FUNCTION_BLOCK basicSubestacao (* Logica unica do QGBT da Subestacao: Masterpact, fonte das barras, planta nos geradores e cargas liberadas *)
  (* Standard: 61499-2 *)
  (* Version 1.3, 04/11/2026, Hidryco, Hidryco, 1.3: comandos do legado REQ_ABRIR_/REQ_FECHAR_1Qx (hmiAbrir/hmiFechar1qx TRUE = mesmo comando do hmiCmdDisjuntor, mesmas permissoes e pulso; FALSE nao faz nada). 1.2: anel - disjuntor com fechamento pendente conta como fechado e o pulso de fechar e cortado se o anel deixar de ter um aberto (nunca as duas QTAM em paralelo). 1.1: comandos de abrir/fechar dos Masterpact 1Q1/1Q0/1Q2 com intertravamentos e aviso de sem resposta; reservas no unifilar. 1.0: QGBT 440 V com 2 QTAM (AGC 150), 1Q1/1Q0/1Q2 e cargas liberadas no gerador *)
  PACKAGE Hidryco.HidrycoLib;
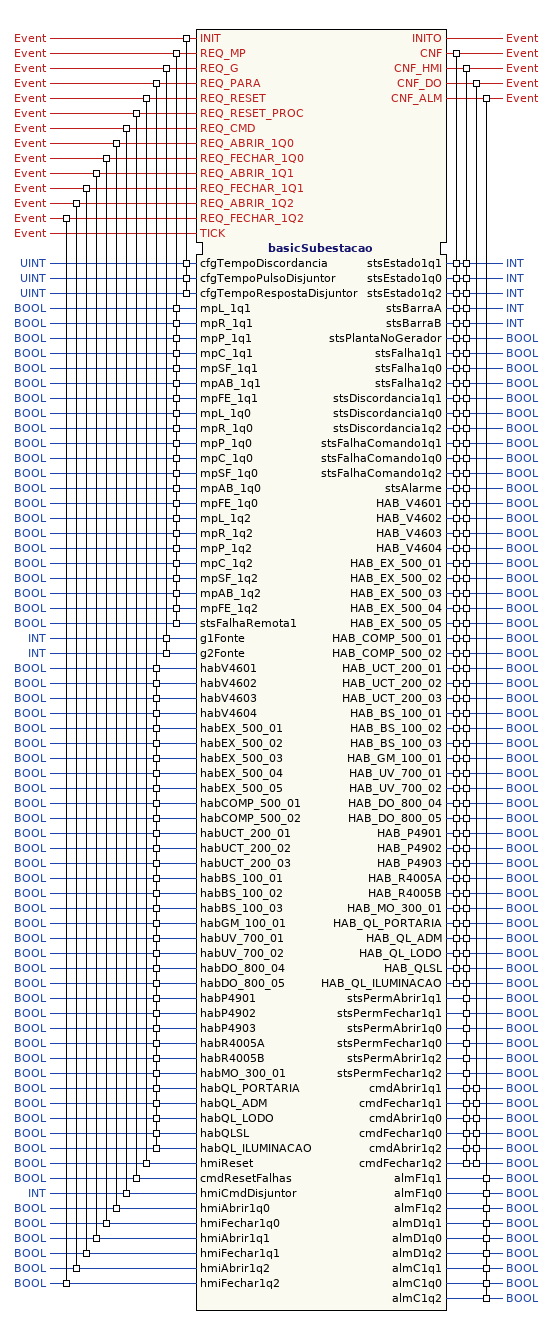
  EVENT_INPUT
    INIT WITH cfgTempoDiscordancia, cfgTempoPulsoDisjuntor, cfgTempoRespostaDisjuntor; (* Inicializacao *)
    REQ_MP WITH mpL_1q1, mpR_1q1, mpP_1q1, mpC_1q1, mpSF_1q1, mpAB_1q1, mpFE_1q1, mpL_1q0, mpR_1q0, mpP_1q0, mpC_1q0, mpSF_1q0, mpAB_1q0, mpFE_1q0, mpL_1q2, mpR_1q2, mpP_1q2, mpC_1q2, mpSF_1q2, mpAB_1q2, mpFE_1q2, stsFalhaRemota1; (* Sinais dos Masterpact e da remota 1 *)
    REQ_G WITH g1Fonte, g2Fonte; (* Estado das QTAM (geradores) *)
    REQ_PARA WITH habV4601, habV4602, habV4603, habV4604, habEX_500_01, habEX_500_02, habEX_500_03, habEX_500_04, habEX_500_05, habCOMP_500_01, habCOMP_500_02, habUCT_200_01, habUCT_200_02, habUCT_200_03, habBS_100_01, habBS_100_02, habBS_100_03, habGM_100_01, habUV_700_01, habUV_700_02, habDO_800_04, habDO_800_05, habP4901, habP4902, habP4903, habR4005A, habR4005B, habMO_300_01, habQL_PORTARIA, habQL_ADM, habQL_LODO, habQLSL, habQL_ILUMINACAO; (* Cargas liberadas no gerador (persistentes) *)
    REQ_RESET WITH hmiReset; (* Reconhecimento pela IHM *)
    REQ_RESET_PROC WITH cmdResetFalhas; (* Reconhecimento pelo processo *)
    REQ_CMD WITH hmiCmdDisjuntor; (* Comando da IHM para os Masterpact *)
    REQ_ABRIR_1Q0 WITH hmiAbrir1q0; (* IHM (legado): ABRIR_1Q0 *)
    REQ_FECHAR_1Q0 WITH hmiFechar1q0; (* IHM (legado): FECHAR_1Q0 *)
    REQ_ABRIR_1Q1 WITH hmiAbrir1q1; (* IHM (legado): ABRIR_1Q1 *)
    REQ_FECHAR_1Q1 WITH hmiFechar1q1; (* IHM (legado): FECHAR_1Q1 *)
    REQ_ABRIR_1Q2 WITH hmiAbrir1q2; (* IHM (legado): ABRIR_1Q2 *)
    REQ_FECHAR_1Q2 WITH hmiFechar1q2; (* IHM (legado): FECHAR_1Q2 *)
    TICK; (* Base de tempo de 1 s *)
  END_EVENT
  EVENT_OUTPUT
    INITO; (* Inicializacao concluida *)
    CNF WITH stsEstado1q1, stsEstado1q0, stsEstado1q2, stsBarraA, stsBarraB, stsPlantaNoGerador, stsFalha1q1, stsFalha1q0, stsFalha1q2, stsDiscordancia1q1, stsDiscordancia1q0, stsDiscordancia1q2, stsFalhaComando1q1, stsFalhaComando1q0, stsFalhaComando1q2, stsAlarme, HAB_V4601, HAB_V4602, HAB_V4603, HAB_V4604, HAB_EX_500_01, HAB_EX_500_02, HAB_EX_500_03, HAB_EX_500_04, HAB_EX_500_05, HAB_COMP_500_01, HAB_COMP_500_02, HAB_UCT_200_01, HAB_UCT_200_02, HAB_UCT_200_03, HAB_BS_100_01, HAB_BS_100_02, HAB_BS_100_03, HAB_GM_100_01, HAB_UV_700_01, HAB_UV_700_02, HAB_DO_800_04, HAB_DO_800_05, HAB_P4901, HAB_P4902, HAB_P4903, HAB_R4005A, HAB_R4005B, HAB_MO_300_01, HAB_QL_PORTARIA, HAB_QL_ADM, HAB_QL_LODO, HAB_QLSL, HAB_QL_ILUMINACAO; (* Estados e cargas liberadas (na mudanca) *)
    CNF_HMI WITH stsEstado1q1, stsEstado1q0, stsEstado1q2, stsBarraA, stsBarraB, stsPlantaNoGerador, stsFalha1q1, stsFalha1q0, stsFalha1q2, stsDiscordancia1q1, stsDiscordancia1q0, stsDiscordancia1q2, stsFalhaComando1q1, stsFalhaComando1q0, stsFalhaComando1q2, stsAlarme, HAB_V4601, HAB_V4602, HAB_V4603, HAB_V4604, HAB_EX_500_01, HAB_EX_500_02, HAB_EX_500_03, HAB_EX_500_04, HAB_EX_500_05, HAB_COMP_500_01, HAB_COMP_500_02, HAB_UCT_200_01, HAB_UCT_200_02, HAB_UCT_200_03, HAB_BS_100_01, HAB_BS_100_02, HAB_BS_100_03, HAB_GM_100_01, HAB_UV_700_01, HAB_UV_700_02, HAB_DO_800_04, HAB_DO_800_05, HAB_P4901, HAB_P4902, HAB_P4903, HAB_R4005A, HAB_R4005B, HAB_MO_300_01, HAB_QL_PORTARIA, HAB_QL_ADM, HAB_QL_LODO, HAB_QLSL, HAB_QL_ILUMINACAO, stsPermAbrir1q1, stsPermFechar1q1, stsPermAbrir1q0, stsPermFechar1q0, stsPermAbrir1q2, stsPermFechar1q2, cmdAbrir1q1, cmdFechar1q1, cmdAbrir1q0, cmdFechar1q0, cmdAbrir1q2, cmdFechar1q2; (* Status para a IHM (na mudanca) *)
    CNF_DO WITH cmdAbrir1q1, cmdFechar1q1, cmdAbrir1q0, cmdFechar1q0, cmdAbrir1q2, cmdFechar1q2; (* Comandos dos Masterpact para o A8 da remota 1 (na mudanca) *)
    CNF_ALM WITH almF1q1, almF1q0, almF1q2, almD1q1, almD1q0, almD1q2, almC1q1, almC1q0, almC1q2; (* Alarmes para os ALARM_BIT (na mudanca) *)
  END_EVENT
  VAR_INPUT
    cfgTempoDiscordancia : UINT := 5; (* Tempo (s) com aberto/fechado discordantes para o aviso de posicao indefinida *)
    cfgTempoPulsoDisjuntor : UINT := 1; (* Tempo (s) do pulso de abrir/fechar dos Masterpact (o pulso acaba antes se o disjuntor mudar de estado) *)
    cfgTempoRespostaDisjuntor : UINT := 5; (* Tempo (s) para o Masterpact mudar de estado depois do comando (senao: aviso de sem resposta) *)
    mpL_1q1 : BOOL; (* Local 1Q1 *)
    mpR_1q1 : BOOL; (* Remoto 1Q1 *)
    mpP_1q1 : BOOL; (* Pronto para fechar 1Q1 *)
    mpC_1q1 : BOOL; (* Mola carregada 1Q1 *)
    mpSF_1q1 : BOOL; (* Sem falha 1Q1 *)
    mpAB_1q1 : BOOL; (* Aberto 1Q1 *)
    mpFE_1q1 : BOOL; (* Fechado 1Q1 *)
    mpL_1q0 : BOOL; (* Local 1Q0 *)
    mpR_1q0 : BOOL; (* Remoto 1Q0 *)
    mpP_1q0 : BOOL; (* Pronto para fechar 1Q0 *)
    mpC_1q0 : BOOL; (* Mola carregada 1Q0 *)
    mpSF_1q0 : BOOL; (* Sem falha 1Q0 *)
    mpAB_1q0 : BOOL; (* Aberto 1Q0 *)
    mpFE_1q0 : BOOL; (* Fechado 1Q0 *)
    mpL_1q2 : BOOL; (* Local 1Q2 *)
    mpR_1q2 : BOOL; (* Remoto 1Q2 *)
    mpP_1q2 : BOOL; (* Pronto para fechar 1Q2 *)
    mpC_1q2 : BOOL; (* Mola carregada 1Q2 *)
    mpSF_1q2 : BOOL; (* Sem falha 1Q2 *)
    mpAB_1q2 : BOOL; (* Aberto 1Q2 *)
    mpFE_1q2 : BOOL; (* Fechado 1Q2 *)
    stsFalhaRemota1 : BOOL; (* Falha de comunicacao com a remota 1 *)
    g1Fonte : INT; (* G1 (QTAM 2): fonte da saida (0 sem, 1 rede, 2 gerador, 3 indefinida) *)
    g2Fonte : INT; (* G2 (QTAM 1): fonte da saida *)
    habV4601 : BOOL; (* IHM: V4601 - Soprador 01 liberado no gerador *)
    habV4602 : BOOL; (* IHM: V4602 - Soprador 02 liberado no gerador *)
    habV4603 : BOOL; (* IHM: V4603 - Soprador 03 liberado no gerador *)
    habV4604 : BOOL; (* IHM: V4604 - Soprador 04 liberado no gerador *)
    habEX_500_01 : BOOL; (* IHM: 500-EX-01 - Exaustor 01 liberado no gerador *)
    habEX_500_02 : BOOL; (* IHM: 500-EX-02 - Exaustor 02 liberado no gerador *)
    habEX_500_03 : BOOL; (* IHM: 500-EX-03 - Exaustor 03 liberado no gerador *)
    habEX_500_04 : BOOL; (* IHM: 500-EX-04 - Exaustor 04 liberado no gerador *)
    habEX_500_05 : BOOL; (* IHM: 500-EX-05 - Exaustor 05 liberado no gerador *)
    habCOMP_500_01 : BOOL; (* IHM: 500-COMP-01 - Compressor 01 liberado no gerador *)
    habCOMP_500_02 : BOOL; (* IHM: 500-COMP-02 - Compressor 02 liberado no gerador *)
    habUCT_200_01 : BOOL; (* IHM: 200-UCT-01 - Unid. compacta 01 liberado no gerador *)
    habUCT_200_02 : BOOL; (* IHM: 200-UCT-02 - Unid. compacta 02 liberado no gerador *)
    habUCT_200_03 : BOOL; (* IHM: 200-UCT-03 - Unid. compacta 03 liberado no gerador *)
    habBS_100_01 : BOOL; (* IHM: 100-BS-01 - Bomba 01 liberado no gerador *)
    habBS_100_02 : BOOL; (* IHM: 100-BS-02 - Bomba 02 liberado no gerador *)
    habBS_100_03 : BOOL; (* IHM: 100-BS-03 - Bomba 03 liberado no gerador *)
    habGM_100_01 : BOOL; (* IHM: 100-GM-01 - Grade mecanizada liberado no gerador *)
    habUV_700_01 : BOOL; (* IHM: 700-UV-01 - Sistema UV 01 liberado no gerador *)
    habUV_700_02 : BOOL; (* IHM: 700-UV-02 - Sistema UV 02 liberado no gerador *)
    habDO_800_04 : BOOL; (* IHM: 800-DO-04 - Bomba dosadora 04 liberado no gerador *)
    habDO_800_05 : BOOL; (* IHM: 800-DO-05 - Bomba dosadora 05 liberado no gerador *)
    habP4901 : BOOL; (* IHM: P4901 - Bomba submersível 01 liberado no gerador *)
    habP4902 : BOOL; (* IHM: P4902 - Bomba submersível 02 liberado no gerador *)
    habP4903 : BOOL; (* IHM: P4903 - Bomba submersível 03 liberado no gerador *)
    habR4005A : BOOL; (* IHM: R4005A - Bomba horizontal A liberado no gerador *)
    habR4005B : BOOL; (* IHM: R4005B - Bomba horizontal B liberado no gerador *)
    habMO_300_01 : BOOL; (* IHM: 300-MO-01 - Misturador 01 liberado no gerador *)
    habQL_PORTARIA : BOOL; (* IHM: QL Portaria liberado no gerador *)
    habQL_ADM : BOOL; (* IHM: QL Administração liberado no gerador *)
    habQL_LODO : BOOL; (* IHM: QL Lodo liberado no gerador *)
    habQLSL : BOOL; (* IHM: QL Sala de quadros liberado no gerador *)
    habQL_ILUMINACAO : BOOL; (* IHM: QL Iluminação externa liberado no gerador *)
    hmiReset : BOOL; (* IHM: reconhecimento *)
    cmdResetFalhas : BOOL; (* Processo: reconhecimento (com E_RESET_FALHAS) *)
    hmiCmdDisjuntor : INT; (* IHM: 1 abrir 1Q1, 2 fechar 1Q1, 3 abrir 1Q0, 4 fechar 1Q0, 5 abrir 1Q2, 6 fechar 1Q2 *)
    hmiAbrir1q0 : BOOL; (* IHM (legado): ABRIR_1Q0, TRUE = executa *)
    hmiFechar1q0 : BOOL; (* IHM (legado): FECHAR_1Q0, TRUE = executa *)
    hmiAbrir1q1 : BOOL; (* IHM (legado): ABRIR_1Q1, TRUE = executa *)
    hmiFechar1q1 : BOOL; (* IHM (legado): FECHAR_1Q1, TRUE = executa *)
    hmiAbrir1q2 : BOOL; (* IHM (legado): ABRIR_1Q2, TRUE = executa *)
    hmiFechar1q2 : BOOL; (* IHM (legado): FECHAR_1Q2, TRUE = executa *)
  END_VAR
  VAR_OUTPUT
    stsEstado1q1 : INT; (* Disjuntor 1Q1: 0 indefinido (sem comunicacao), 1 aberto, 2 fechado, 3 discordante *)
    stsEstado1q0 : INT; (* Disjuntor 1Q0: 0 indefinido (sem comunicacao), 1 aberto, 2 fechado, 3 discordante *)
    stsEstado1q2 : INT; (* Disjuntor 1Q2: 0 indefinido (sem comunicacao), 1 aberto, 2 fechado, 3 discordante *)
    stsBarraA : INT; (* Fonte da barra A (1Q1): 0 sem alimentacao, 1 rede, 2 gerador, 3 indefinida *)
    stsBarraB : INT; (* Fonte da barra B (1Q2): 0 sem alimentacao, 1 rede, 2 gerador, 3 indefinida *)
    stsPlantaNoGerador : BOOL; (* Alguma QTAM com o disjuntor do gerador fechado (planta nos geradores) *)
    stsFalha1q1 : BOOL; (* Disjuntor 1Q1 em falha (desarmado) *)
    stsFalha1q0 : BOOL; (* Disjuntor 1Q0 em falha (desarmado) *)
    stsFalha1q2 : BOOL; (* Disjuntor 1Q2 em falha (desarmado) *)
    stsDiscordancia1q1 : BOOL; (* Disjuntor 1Q1: posição indefinida (aberto e fechado discordantes) *)
    stsDiscordancia1q0 : BOOL; (* Disjuntor 1Q0: posição indefinida (aberto e fechado discordantes) *)
    stsDiscordancia1q2 : BOOL; (* Disjuntor 1Q2: posição indefinida (aberto e fechado discordantes) *)
    stsFalhaComando1q1 : BOOL; (* Disjuntor 1Q1 não respondeu ao comando de abrir/fechar *)
    stsFalhaComando1q0 : BOOL; (* Disjuntor 1Q0 não respondeu ao comando de abrir/fechar *)
    stsFalhaComando1q2 : BOOL; (* Disjuntor 1Q2 não respondeu ao comando de abrir/fechar *)
    stsAlarme : BOOL; (* Algum alarme do QGBT *)
    HAB_V4601 : BOOL; (* V4601 - Soprador 01 liberado para operar com a planta nos geradores *)
    HAB_V4602 : BOOL; (* V4602 - Soprador 02 liberado para operar com a planta nos geradores *)
    HAB_V4603 : BOOL; (* V4603 - Soprador 03 liberado para operar com a planta nos geradores *)
    HAB_V4604 : BOOL; (* V4604 - Soprador 04 liberado para operar com a planta nos geradores *)
    HAB_EX_500_01 : BOOL; (* 500-EX-01 - Exaustor 01 liberado para operar com a planta nos geradores *)
    HAB_EX_500_02 : BOOL; (* 500-EX-02 - Exaustor 02 liberado para operar com a planta nos geradores *)
    HAB_EX_500_03 : BOOL; (* 500-EX-03 - Exaustor 03 liberado para operar com a planta nos geradores *)
    HAB_EX_500_04 : BOOL; (* 500-EX-04 - Exaustor 04 liberado para operar com a planta nos geradores *)
    HAB_EX_500_05 : BOOL; (* 500-EX-05 - Exaustor 05 liberado para operar com a planta nos geradores *)
    HAB_COMP_500_01 : BOOL; (* 500-COMP-01 - Compressor 01 liberado para operar com a planta nos geradores *)
    HAB_COMP_500_02 : BOOL; (* 500-COMP-02 - Compressor 02 liberado para operar com a planta nos geradores *)
    HAB_UCT_200_01 : BOOL; (* 200-UCT-01 - Unid. compacta 01 liberado para operar com a planta nos geradores *)
    HAB_UCT_200_02 : BOOL; (* 200-UCT-02 - Unid. compacta 02 liberado para operar com a planta nos geradores *)
    HAB_UCT_200_03 : BOOL; (* 200-UCT-03 - Unid. compacta 03 liberado para operar com a planta nos geradores *)
    HAB_BS_100_01 : BOOL; (* 100-BS-01 - Bomba 01 liberado para operar com a planta nos geradores *)
    HAB_BS_100_02 : BOOL; (* 100-BS-02 - Bomba 02 liberado para operar com a planta nos geradores *)
    HAB_BS_100_03 : BOOL; (* 100-BS-03 - Bomba 03 liberado para operar com a planta nos geradores *)
    HAB_GM_100_01 : BOOL; (* 100-GM-01 - Grade mecanizada liberado para operar com a planta nos geradores *)
    HAB_UV_700_01 : BOOL; (* 700-UV-01 - Sistema UV 01 liberado para operar com a planta nos geradores *)
    HAB_UV_700_02 : BOOL; (* 700-UV-02 - Sistema UV 02 liberado para operar com a planta nos geradores *)
    HAB_DO_800_04 : BOOL; (* 800-DO-04 - Bomba dosadora 04 liberado para operar com a planta nos geradores *)
    HAB_DO_800_05 : BOOL; (* 800-DO-05 - Bomba dosadora 05 liberado para operar com a planta nos geradores *)
    HAB_P4901 : BOOL; (* P4901 - Bomba submersível 01 liberado para operar com a planta nos geradores *)
    HAB_P4902 : BOOL; (* P4902 - Bomba submersível 02 liberado para operar com a planta nos geradores *)
    HAB_P4903 : BOOL; (* P4903 - Bomba submersível 03 liberado para operar com a planta nos geradores *)
    HAB_R4005A : BOOL; (* R4005A - Bomba horizontal A liberado para operar com a planta nos geradores *)
    HAB_R4005B : BOOL; (* R4005B - Bomba horizontal B liberado para operar com a planta nos geradores *)
    HAB_MO_300_01 : BOOL; (* 300-MO-01 - Misturador 01 liberado para operar com a planta nos geradores *)
    HAB_QL_PORTARIA : BOOL; (* QL Portaria liberado para operar com a planta nos geradores *)
    HAB_QL_ADM : BOOL; (* QL Administração liberado para operar com a planta nos geradores *)
    HAB_QL_LODO : BOOL; (* QL Lodo liberado para operar com a planta nos geradores *)
    HAB_QLSL : BOOL; (* QL Sala de quadros liberado para operar com a planta nos geradores *)
    HAB_QL_ILUMINACAO : BOOL; (* QL Iluminação externa liberado para operar com a planta nos geradores *)
    stsPermAbrir1q1 : BOOL; (* IHM: abrir o 1Q1 permitido *)
    stsPermFechar1q1 : BOOL; (* IHM: fechar o 1Q1 permitido *)
    stsPermAbrir1q0 : BOOL; (* IHM: abrir o 1Q0 permitido *)
    stsPermFechar1q0 : BOOL; (* IHM: fechar o 1Q0 permitido *)
    stsPermAbrir1q2 : BOOL; (* IHM: abrir o 1Q2 permitido *)
    stsPermFechar1q2 : BOOL; (* IHM: fechar o 1Q2 permitido *)
    cmdAbrir1q1 : BOOL; (* Pulso de abrir o 1Q1 (bobina MX) *)
    cmdFechar1q1 : BOOL; (* Pulso de fechar o 1Q1 (bobina XF) *)
    cmdAbrir1q0 : BOOL; (* Pulso de abrir o 1Q0 (bobina MX) *)
    cmdFechar1q0 : BOOL; (* Pulso de fechar o 1Q0 (bobina XF) *)
    cmdAbrir1q2 : BOOL; (* Pulso de abrir o 1Q2 (bobina MX) *)
    cmdFechar1q2 : BOOL; (* Pulso de fechar o 1Q2 (bobina XF) *)
    almF1q1 : BOOL; (* ALARM_BIT Disjuntor 1Q1 em falha (desarmado) *)
    almF1q0 : BOOL; (* ALARM_BIT Disjuntor 1Q0 em falha (desarmado) *)
    almF1q2 : BOOL; (* ALARM_BIT Disjuntor 1Q2 em falha (desarmado) *)
    almD1q1 : BOOL; (* ALARM_BIT Disjuntor 1Q1: posição indefinida (aberto e fechado discordantes) *)
    almD1q0 : BOOL; (* ALARM_BIT Disjuntor 1Q0: posição indefinida (aberto e fechado discordantes) *)
    almD1q2 : BOOL; (* ALARM_BIT Disjuntor 1Q2: posição indefinida (aberto e fechado discordantes) *)
    almC1q1 : BOOL; (* ALARM_BIT Disjuntor 1Q1 não respondeu ao comando de abrir/fechar *)
    almC1q0 : BOOL; (* ALARM_BIT Disjuntor 1Q0 não respondeu ao comando de abrir/fechar *)
    almC1q2 : BOOL; (* ALARM_BIT Disjuntor 1Q2 não respondeu ao comando de abrir/fechar *)
  END_VAR
  VAR
    cmdDj : INT; (* Comando do disjuntor deste ciclo (hmiCmdDisjuntor ou comando do legado) *)
    initDone : BOOL;
    initPass : BOOL;
    bMudou : BOOL;
    u1q1 : UDINT; (* Segundos com aberto/fechado discordantes *)
    u1q0 : UDINT; (* Segundos com aberto/fechado discordantes *)
    u1q2 : UDINT; (* Segundos com aberto/fechado discordantes *)
    e1q1 : INT;
    e1q0 : INT;
    e1q2 : INT;
    wSts : DWORD;
    oldSts : DWORD := 16#FFFFFFFF;
    wHab : DWORD;
    oldHab : DWORD := 16#FFFFFFFF;
    wHab2 : DWORD;
    oldHab2 : DWORD := 16#FFFFFFFF;
    wAlm : WORD;
    oldAlm : WORD := 16#FFFF;
    wPerm : WORD;
    oldPerm : WORD := 16#FFFF;
    wDo : WORD;
    oldDo : WORD := 16#FFFF;
    o_stsEstado1q1 : INT := -1;
    o_stsEstado1q0 : INT := -1;
    o_stsEstado1q2 : INT := -1;
    o_stsBarraA : INT := -1;
    o_stsBarraB : INT := -1;
    tA1q1 : UINT; (* Pulso de abrir restante (s) *)
    tF1q1 : UINT; (* Pulso de fechar restante (s) *)
    uR1q1 : UINT; (* Tempo restante para a resposta (s) *)
    tA1q0 : UINT; (* Pulso de abrir restante (s) *)
    tF1q0 : UINT; (* Pulso de fechar restante (s) *)
    uR1q0 : UINT; (* Tempo restante para a resposta (s) *)
    tA1q2 : UINT; (* Pulso de abrir restante (s) *)
    tF1q2 : UINT; (* Pulso de fechar restante (s) *)
    uR1q2 : UINT; (* Tempo restante para a resposta (s) *)
    alvo1q1 : INT; (* Estado esperado depois do comando (0 nenhum, 1 aberto, 2 fechado) *)
    alvo1q0 : INT; (* Estado esperado depois do comando (0 nenhum, 1 aberto, 2 fechado) *)
    alvo1q2 : INT; (* Estado esperado depois do comando (0 nenhum, 1 aberto, 2 fechado) *)
  END_VAR
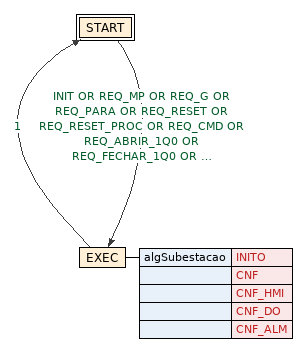
  EC_STATES
    START; (* Estado inicial *)
    EXEC : algSubestacao -> INITO, -> CNF, -> CNF_HMI, -> CNF_DO, -> CNF_ALM; (* Executa a logica; o algoritmo decide quais eventos saem *)
  END_STATES
  EC_TRANSITIONS
    START TO EXEC := INIT OR REQ_MP OR REQ_G OR REQ_PARA OR REQ_RESET OR REQ_RESET_PROC OR REQ_CMD OR REQ_ABRIR_1Q0 OR REQ_FECHAR_1Q0 OR REQ_ABRIR_1Q1 OR REQ_FECHAR_1Q1 OR REQ_ABRIR_1Q2 OR REQ_FECHAR_1Q2 OR TICK;
    EXEC TO START := 1;
  END_TRANSITIONS
  ALGORITHM algSubestacao IN ST: (* Logica completa do QGBT (um unico algoritmo) *)
(* =====================================================================
   basicSubestacao v1.1 - QGBT 440 V da ETE Tijuco Preto
   QTAM 1 (G2) -> 1Q1 -> barra A; QTAM 2 (G1) -> 1Q2 -> barra B; 1Q0 acopla.
   - Masterpact: 2 fechado, 1 aberto, 3 aberto/fechado discordantes,
     0 indefinido (remota 1 sem comunicacao); aviso de discordancia apos
     cfgTempoDiscordancia s; alarme de falha com "sem falha" = FALSE;
   - fonte de cada barra pelo seu Masterpact ou pelo acoplamento 1Q0;
   - planta nos geradores = alguma QTAM com o disjuntor do gerador fechado
     (vale mesmo com a remota 1 sem comunicacao);
   - cargas liberadas no gerador: escolha do operador (persistente), saidas
     HAB_* para os CATs de processo (geradorHabilita);
   - v1.1: comandos de abrir/fechar dos Masterpact com intertravamentos.
   ===================================================================== *)

INITO   := FALSE;
CNF     := FALSE;
CNF_HMI := FALSE;
CNF_DO  := FALSE;
CNF_ALM := FALSE;
IF INIT THEN
    initDone := TRUE;
    initPass := TRUE;
    INITO    := TRUE;
END_IF;
IF NOT initDone THEN
    RETURN;
END_IF;

(* ---- 1Q1 ---- *)
IF stsFalhaRemota1 THEN
    e1q1 := 0;
ELSIF mpAB_1q1 AND NOT mpFE_1q1 THEN
    e1q1 := 1;
ELSIF mpFE_1q1 AND NOT mpAB_1q1 THEN
    e1q1 := 2;
ELSE
    e1q1 := 3;
END_IF;
IF e1q1 = 3 THEN
    IF TICK AND u1q1 < UINT_TO_UDINT(cfgTempoDiscordancia) THEN
        u1q1 := u1q1 + 1;
    END_IF;
ELSE
    u1q1 := 0;
END_IF;
stsEstado1q1 := e1q1;
stsDiscordancia1q1 := e1q1 = 3 AND u1q1 >= UINT_TO_UDINT(cfgTempoDiscordancia);
stsFalha1q1 := NOT stsFalhaRemota1 AND NOT mpSF_1q1;

(* ---- 1Q0 ---- *)
IF stsFalhaRemota1 THEN
    e1q0 := 0;
ELSIF mpAB_1q0 AND NOT mpFE_1q0 THEN
    e1q0 := 1;
ELSIF mpFE_1q0 AND NOT mpAB_1q0 THEN
    e1q0 := 2;
ELSE
    e1q0 := 3;
END_IF;
IF e1q0 = 3 THEN
    IF TICK AND u1q0 < UINT_TO_UDINT(cfgTempoDiscordancia) THEN
        u1q0 := u1q0 + 1;
    END_IF;
ELSE
    u1q0 := 0;
END_IF;
stsEstado1q0 := e1q0;
stsDiscordancia1q0 := e1q0 = 3 AND u1q0 >= UINT_TO_UDINT(cfgTempoDiscordancia);
stsFalha1q0 := NOT stsFalhaRemota1 AND NOT mpSF_1q0;

(* ---- 1Q2 ---- *)
IF stsFalhaRemota1 THEN
    e1q2 := 0;
ELSIF mpAB_1q2 AND NOT mpFE_1q2 THEN
    e1q2 := 1;
ELSIF mpFE_1q2 AND NOT mpAB_1q2 THEN
    e1q2 := 2;
ELSE
    e1q2 := 3;
END_IF;
IF e1q2 = 3 THEN
    IF TICK AND u1q2 < UINT_TO_UDINT(cfgTempoDiscordancia) THEN
        u1q2 := u1q2 + 1;
    END_IF;
ELSE
    u1q2 := 0;
END_IF;
stsEstado1q2 := e1q2;
stsDiscordancia1q2 := e1q2 = 3 AND u1q2 >= UINT_TO_UDINT(cfgTempoDiscordancia);
stsFalha1q2 := NOT stsFalhaRemota1 AND NOT mpSF_1q2;

(* ---- fonte das barras: 0 sem alimentacao, 1 rede, 2 gerador, 3 indefinida ---- *)
IF e1q1 = 2 THEN
    stsBarraA := g2Fonte;
ELSIF e1q1 = 1 AND e1q0 = 2 AND e1q2 = 2 THEN
    stsBarraA := g1Fonte;
ELSIF e1q1 = 1 AND (e1q0 = 1 OR e1q2 = 1) THEN
    stsBarraA := 0;
ELSE
    stsBarraA := 3;
END_IF;
IF e1q2 = 2 THEN
    stsBarraB := g1Fonte;
ELSIF e1q2 = 1 AND e1q0 = 2 AND e1q1 = 2 THEN
    stsBarraB := g2Fonte;
ELSIF e1q2 = 1 AND (e1q0 = 1 OR e1q1 = 1) THEN
    stsBarraB := 0;
ELSE
    stsBarraB := 3;
END_IF;
stsPlantaNoGerador := g1Fonte = 2 OR g2Fonte = 2;

(* ---- cargas liberadas no gerador (escolha do operador) ---- *)
HAB_V4601 := habV4601;
HAB_V4602 := habV4602;
HAB_V4603 := habV4603;
HAB_V4604 := habV4604;
HAB_EX_500_01 := habEX_500_01;
HAB_EX_500_02 := habEX_500_02;
HAB_EX_500_03 := habEX_500_03;
HAB_EX_500_04 := habEX_500_04;
HAB_EX_500_05 := habEX_500_05;
HAB_COMP_500_01 := habCOMP_500_01;
HAB_COMP_500_02 := habCOMP_500_02;
HAB_UCT_200_01 := habUCT_200_01;
HAB_UCT_200_02 := habUCT_200_02;
HAB_UCT_200_03 := habUCT_200_03;
HAB_BS_100_01 := habBS_100_01;
HAB_BS_100_02 := habBS_100_02;
HAB_BS_100_03 := habBS_100_03;
HAB_GM_100_01 := habGM_100_01;
HAB_UV_700_01 := habUV_700_01;
HAB_UV_700_02 := habUV_700_02;
HAB_DO_800_04 := habDO_800_04;
HAB_DO_800_05 := habDO_800_05;
HAB_P4901 := habP4901;
HAB_P4902 := habP4902;
HAB_P4903 := habP4903;
HAB_R4005A := habR4005A;
HAB_R4005B := habR4005B;
HAB_MO_300_01 := habMO_300_01;
HAB_QL_PORTARIA := habQL_PORTARIA;
HAB_QL_ADM := habQL_ADM;
HAB_QL_LODO := habQL_LODO;
HAB_QLSL := habQLSL;
HAB_QL_ILUMINACAO := habQL_ILUMINACAO;

(* ---- comandos dos Masterpact (IHM) ----
   abrir: remota OK, fechado, em remoto (nao local);
   fechar: remota OK, aberto, remoto, pronto para fechar, mola carregada, sem falha
           e sem fechar o anel: 1Q1 e 1Q2 so com o 1Q0 ou o outro aberto;
           1Q0 so com o 1Q1 ou o 1Q2 aberto (nunca as duas QTAM em paralelo);
           disjuntor com fechamento pendente conta como fechado; pulso de fechar e cortado
           se o anel deixar de ter um disjuntor aberto;
   pulso de cfgTempoPulsoDisjuntor s (acaba antes se o disjuntor mudar);
   sem mudanca em cfgTempoRespostaDisjuntor s: aviso de sem resposta. *)
stsPermAbrir1q1 := NOT stsFalhaRemota1 AND e1q1 = 2 AND mpR_1q1 AND NOT mpL_1q1;
stsPermFechar1q1 := NOT stsFalhaRemota1 AND e1q1 = 1 AND mpR_1q1 AND NOT mpL_1q1 AND mpP_1q1 AND mpC_1q1 AND mpSF_1q1 AND ((e1q0 = 1 AND alvo1q0 <> 2) OR (e1q2 = 1 AND alvo1q2 <> 2));
stsPermAbrir1q0 := NOT stsFalhaRemota1 AND e1q0 = 2 AND mpR_1q0 AND NOT mpL_1q0;
stsPermFechar1q0 := NOT stsFalhaRemota1 AND e1q0 = 1 AND mpR_1q0 AND NOT mpL_1q0 AND mpP_1q0 AND mpC_1q0 AND mpSF_1q0 AND ((e1q1 = 1 AND alvo1q1 <> 2) OR (e1q2 = 1 AND alvo1q2 <> 2));
stsPermAbrir1q2 := NOT stsFalhaRemota1 AND e1q2 = 2 AND mpR_1q2 AND NOT mpL_1q2;
stsPermFechar1q2 := NOT stsFalhaRemota1 AND e1q2 = 1 AND mpR_1q2 AND NOT mpL_1q2 AND mpP_1q2 AND mpC_1q2 AND mpSF_1q2 AND ((e1q0 = 1 AND alvo1q0 <> 2) OR (e1q1 = 1 AND alvo1q1 <> 2));
cmdDj := 0;
IF REQ_CMD THEN
    cmdDj := hmiCmdDisjuntor;
END_IF;
(* comandos do legado: TRUE executa; FALSE nao faz nada *)
IF REQ_ABRIR_1Q0 AND hmiAbrir1q0 THEN
    cmdDj := 3;
END_IF;
IF REQ_FECHAR_1Q0 AND hmiFechar1q0 THEN
    cmdDj := 4;
END_IF;
IF REQ_ABRIR_1Q1 AND hmiAbrir1q1 THEN
    cmdDj := 1;
END_IF;
IF REQ_FECHAR_1Q1 AND hmiFechar1q1 THEN
    cmdDj := 2;
END_IF;
IF REQ_ABRIR_1Q2 AND hmiAbrir1q2 THEN
    cmdDj := 5;
END_IF;
IF REQ_FECHAR_1Q2 AND hmiFechar1q2 THEN
    cmdDj := 6;
END_IF;
IF cmdDj <> 0 THEN
    IF cmdDj = 1 AND stsPermAbrir1q1 THEN
        tF1q1 := 0;
        tA1q1 := cfgTempoPulsoDisjuntor + 1;
        alvo1q1 := 1;
        uR1q1 := cfgTempoRespostaDisjuntor;
        stsFalhaComando1q1 := FALSE;
    ELSIF cmdDj = 2 AND stsPermFechar1q1 THEN
        tA1q1 := 0;
        tF1q1 := cfgTempoPulsoDisjuntor + 1;
        alvo1q1 := 2;
        uR1q1 := cfgTempoRespostaDisjuntor;
        stsFalhaComando1q1 := FALSE;
    ELSIF cmdDj = 3 AND stsPermAbrir1q0 THEN
        tF1q0 := 0;
        tA1q0 := cfgTempoPulsoDisjuntor + 1;
        alvo1q0 := 1;
        uR1q0 := cfgTempoRespostaDisjuntor;
        stsFalhaComando1q0 := FALSE;
    ELSIF cmdDj = 4 AND stsPermFechar1q0 THEN
        tA1q0 := 0;
        tF1q0 := cfgTempoPulsoDisjuntor + 1;
        alvo1q0 := 2;
        uR1q0 := cfgTempoRespostaDisjuntor;
        stsFalhaComando1q0 := FALSE;
    ELSIF cmdDj = 5 AND stsPermAbrir1q2 THEN
        tF1q2 := 0;
        tA1q2 := cfgTempoPulsoDisjuntor + 1;
        alvo1q2 := 1;
        uR1q2 := cfgTempoRespostaDisjuntor;
        stsFalhaComando1q2 := FALSE;
    ELSIF cmdDj = 6 AND stsPermFechar1q2 THEN
        tA1q2 := 0;
        tF1q2 := cfgTempoPulsoDisjuntor + 1;
        alvo1q2 := 2;
        uR1q2 := cfgTempoRespostaDisjuntor;
        stsFalhaComando1q2 := FALSE;
    END_IF;
END_IF;
IF (REQ_RESET AND hmiReset) OR (REQ_RESET_PROC AND cmdResetFalhas) THEN
    stsFalhaComando1q1 := FALSE;
    stsFalhaComando1q0 := FALSE;
    stsFalhaComando1q2 := FALSE;
END_IF;
IF alvo1q1 > 0 AND e1q1 = alvo1q1 THEN
    tA1q1 := 0;
    tF1q1 := 0;
    alvo1q1 := 0;
    uR1q1 := 0;
END_IF;
IF TICK THEN
    IF tA1q1 > 0 THEN tA1q1 := tA1q1 - 1; END_IF;
    IF tF1q1 > 0 THEN tF1q1 := tF1q1 - 1; END_IF;
    IF alvo1q1 > 0 THEN
        IF uR1q1 > 0 THEN uR1q1 := uR1q1 - 1; END_IF;
        IF uR1q1 = 0 THEN
            stsFalhaComando1q1 := TRUE;
            alvo1q1 := 0;
            tA1q1 := 0;
            tF1q1 := 0;
        END_IF;
    END_IF;
END_IF;
IF stsFalhaRemota1 THEN
    tA1q1 := 0;
    tF1q1 := 0;
END_IF;
cmdAbrir1q1 := tA1q1 > 0;
cmdFechar1q1 := tF1q1 > 0;
IF alvo1q0 > 0 AND e1q0 = alvo1q0 THEN
    tA1q0 := 0;
    tF1q0 := 0;
    alvo1q0 := 0;
    uR1q0 := 0;
END_IF;
IF TICK THEN
    IF tA1q0 > 0 THEN tA1q0 := tA1q0 - 1; END_IF;
    IF tF1q0 > 0 THEN tF1q0 := tF1q0 - 1; END_IF;
    IF alvo1q0 > 0 THEN
        IF uR1q0 > 0 THEN uR1q0 := uR1q0 - 1; END_IF;
        IF uR1q0 = 0 THEN
            stsFalhaComando1q0 := TRUE;
            alvo1q0 := 0;
            tA1q0 := 0;
            tF1q0 := 0;
        END_IF;
    END_IF;
END_IF;
IF stsFalhaRemota1 THEN
    tA1q0 := 0;
    tF1q0 := 0;
END_IF;
cmdAbrir1q0 := tA1q0 > 0;
cmdFechar1q0 := tF1q0 > 0;
IF alvo1q2 > 0 AND e1q2 = alvo1q2 THEN
    tA1q2 := 0;
    tF1q2 := 0;
    alvo1q2 := 0;
    uR1q2 := 0;
END_IF;
IF TICK THEN
    IF tA1q2 > 0 THEN tA1q2 := tA1q2 - 1; END_IF;
    IF tF1q2 > 0 THEN tF1q2 := tF1q2 - 1; END_IF;
    IF alvo1q2 > 0 THEN
        IF uR1q2 > 0 THEN uR1q2 := uR1q2 - 1; END_IF;
        IF uR1q2 = 0 THEN
            stsFalhaComando1q2 := TRUE;
            alvo1q2 := 0;
            tA1q2 := 0;
            tF1q2 := 0;
        END_IF;
    END_IF;
END_IF;
IF stsFalhaRemota1 THEN
    tA1q2 := 0;
    tF1q2 := 0;
END_IF;
cmdAbrir1q2 := tA1q2 > 0;
cmdFechar1q2 := tF1q2 > 0;
(* anel: corta o pulso de fechar se o anel deixou de ter um disjuntor aberto (fechamento no campo durante o pulso) *)
IF tF1q1 > 0 AND NOT ((e1q0 = 1 AND alvo1q0 <> 2) OR (e1q2 = 1 AND alvo1q2 <> 2)) THEN tF1q1 := 0; cmdFechar1q1 := FALSE; END_IF;
IF tF1q0 > 0 AND NOT ((e1q1 = 1 AND alvo1q1 <> 2) OR (e1q2 = 1 AND alvo1q2 <> 2)) THEN tF1q0 := 0; cmdFechar1q0 := FALSE; END_IF;
IF tF1q2 > 0 AND NOT ((e1q0 = 1 AND alvo1q0 <> 2) OR (e1q1 = 1 AND alvo1q1 <> 2)) THEN tF1q2 := 0; cmdFechar1q2 := FALSE; END_IF;

(* ---- alarmes ---- *)
almF1q1 := stsFalha1q1;
almF1q0 := stsFalha1q0;
almF1q2 := stsFalha1q2;
almD1q1 := stsDiscordancia1q1;
almD1q0 := stsDiscordancia1q0;
almD1q2 := stsDiscordancia1q2;
almC1q1 := stsFalhaComando1q1;
almC1q0 := stsFalhaComando1q0;
almC1q2 := stsFalhaComando1q2;
stsAlarme := almF1q1 OR almF1q0 OR almF1q2 OR almD1q1 OR almD1q0 OR almD1q2 OR almC1q1 OR almC1q0 OR almC1q2;

(* ---- eventos so na mudanca ---- *)
bMudou := FALSE;
IF stsEstado1q1 <> o_stsEstado1q1 THEN bMudou := TRUE; o_stsEstado1q1 := stsEstado1q1; END_IF;
IF stsEstado1q0 <> o_stsEstado1q0 THEN bMudou := TRUE; o_stsEstado1q0 := stsEstado1q0; END_IF;
IF stsEstado1q2 <> o_stsEstado1q2 THEN bMudou := TRUE; o_stsEstado1q2 := stsEstado1q2; END_IF;
IF stsBarraA <> o_stsBarraA THEN bMudou := TRUE; o_stsBarraA := stsBarraA; END_IF;
IF stsBarraB <> o_stsBarraB THEN bMudou := TRUE; o_stsBarraB := stsBarraB; END_IF;
wSts := 0;
IF stsPlantaNoGerador THEN wSts := wSts OR 16#00000001; END_IF;
IF stsFalha1q1 THEN wSts := wSts OR 16#00000002; END_IF;
IF stsFalha1q0 THEN wSts := wSts OR 16#00000004; END_IF;
IF stsFalha1q2 THEN wSts := wSts OR 16#00000008; END_IF;
IF stsDiscordancia1q1 THEN wSts := wSts OR 16#00000010; END_IF;
IF stsDiscordancia1q0 THEN wSts := wSts OR 16#00000020; END_IF;
IF stsDiscordancia1q2 THEN wSts := wSts OR 16#00000040; END_IF;
IF stsFalhaComando1q1 THEN wSts := wSts OR 16#00000080; END_IF;
IF stsFalhaComando1q0 THEN wSts := wSts OR 16#00000100; END_IF;
IF stsFalhaComando1q2 THEN wSts := wSts OR 16#00000200; END_IF;
IF stsAlarme THEN wSts := wSts OR 16#00000400; END_IF;
wHab := 0;
wHab2 := 0;
IF HAB_V4601 THEN wHab := wHab OR 16#00000001; END_IF;
IF HAB_V4602 THEN wHab := wHab OR 16#00000002; END_IF;
IF HAB_V4603 THEN wHab := wHab OR 16#00000004; END_IF;
IF HAB_V4604 THEN wHab := wHab OR 16#00000008; END_IF;
IF HAB_EX_500_01 THEN wHab := wHab OR 16#00000010; END_IF;
IF HAB_EX_500_02 THEN wHab := wHab OR 16#00000020; END_IF;
IF HAB_EX_500_03 THEN wHab := wHab OR 16#00000040; END_IF;
IF HAB_EX_500_04 THEN wHab := wHab OR 16#00000080; END_IF;
IF HAB_EX_500_05 THEN wHab := wHab OR 16#00000100; END_IF;
IF HAB_COMP_500_01 THEN wHab := wHab OR 16#00000200; END_IF;
IF HAB_COMP_500_02 THEN wHab := wHab OR 16#00000400; END_IF;
IF HAB_UCT_200_01 THEN wHab := wHab OR 16#00000800; END_IF;
IF HAB_UCT_200_02 THEN wHab := wHab OR 16#00001000; END_IF;
IF HAB_UCT_200_03 THEN wHab := wHab OR 16#00002000; END_IF;
IF HAB_BS_100_01 THEN wHab := wHab OR 16#00004000; END_IF;
IF HAB_BS_100_02 THEN wHab := wHab OR 16#00008000; END_IF;
IF HAB_BS_100_03 THEN wHab := wHab OR 16#00010000; END_IF;
IF HAB_GM_100_01 THEN wHab := wHab OR 16#00020000; END_IF;
IF HAB_UV_700_01 THEN wHab := wHab OR 16#00040000; END_IF;
IF HAB_UV_700_02 THEN wHab := wHab OR 16#00080000; END_IF;
IF HAB_DO_800_04 THEN wHab := wHab OR 16#00100000; END_IF;
IF HAB_DO_800_05 THEN wHab := wHab OR 16#00200000; END_IF;
IF HAB_P4901 THEN wHab := wHab OR 16#00400000; END_IF;
IF HAB_P4902 THEN wHab := wHab OR 16#00800000; END_IF;
IF HAB_P4903 THEN wHab := wHab OR 16#01000000; END_IF;
IF HAB_R4005A THEN wHab := wHab OR 16#02000000; END_IF;
IF HAB_R4005B THEN wHab := wHab OR 16#04000000; END_IF;
IF HAB_MO_300_01 THEN wHab := wHab OR 16#08000000; END_IF;
IF HAB_QL_PORTARIA THEN wHab := wHab OR 16#10000000; END_IF;
IF HAB_QL_ADM THEN wHab := wHab OR 16#20000000; END_IF;
IF HAB_QL_LODO THEN wHab := wHab OR 16#40000000; END_IF;
IF HAB_QLSL THEN wHab := wHab OR 16#80000000; END_IF;
IF HAB_QL_ILUMINACAO THEN wHab2 := wHab2 OR 16#00000001; END_IF;
wAlm := 0;
IF almF1q1 THEN wAlm := wAlm OR 16#0001; END_IF;
IF almF1q0 THEN wAlm := wAlm OR 16#0002; END_IF;
IF almF1q2 THEN wAlm := wAlm OR 16#0004; END_IF;
IF almD1q1 THEN wAlm := wAlm OR 16#0008; END_IF;
IF almD1q0 THEN wAlm := wAlm OR 16#0010; END_IF;
IF almD1q2 THEN wAlm := wAlm OR 16#0020; END_IF;
IF almC1q1 THEN wAlm := wAlm OR 16#0040; END_IF;
IF almC1q0 THEN wAlm := wAlm OR 16#0080; END_IF;
IF almC1q2 THEN wAlm := wAlm OR 16#0100; END_IF;
wPerm := 0;
IF stsPermAbrir1q1 THEN wPerm := wPerm OR 16#0001; END_IF;
IF stsPermFechar1q1 THEN wPerm := wPerm OR 16#0002; END_IF;
IF stsPermAbrir1q0 THEN wPerm := wPerm OR 16#0004; END_IF;
IF stsPermFechar1q0 THEN wPerm := wPerm OR 16#0008; END_IF;
IF stsPermAbrir1q2 THEN wPerm := wPerm OR 16#0010; END_IF;
IF stsPermFechar1q2 THEN wPerm := wPerm OR 16#0020; END_IF;
wDo := 0;
IF cmdAbrir1q1 THEN wDo := wDo OR 16#0001; END_IF;
IF cmdFechar1q1 THEN wDo := wDo OR 16#0002; END_IF;
IF cmdAbrir1q0 THEN wDo := wDo OR 16#0004; END_IF;
IF cmdFechar1q0 THEN wDo := wDo OR 16#0008; END_IF;
IF cmdAbrir1q2 THEN wDo := wDo OR 16#0010; END_IF;
IF cmdFechar1q2 THEN wDo := wDo OR 16#0020; END_IF;
CNF := initPass OR bMudou OR (wSts <> oldSts) OR (wHab <> oldHab) OR (wHab2 <> oldHab2);
CNF_DO := initPass OR (wDo <> oldDo);
CNF_HMI := CNF OR (wPerm <> oldPerm) OR CNF_DO;
CNF_ALM := initPass OR (wAlm <> oldAlm);
oldPerm := wPerm;
oldDo := wDo;
oldSts := wSts;
oldHab := wHab;
oldHab2 := wHab2;
oldAlm := wAlm;
initPass := FALSE;
  END_ALGORITHM
END_FUNCTION_BLOCK
